(* IEC 61131-3 sources: avi-aoi-management/scripts/ai-eval/ngau-nhien/kho/st-ud5-sao-tam-giac/khung/src, 2 files *)

(* ---- KhoaChuyenMach.st ---- *)
FUNCTION_BLOCK KhoaChuyenMach
VAR_INPUT
    YC_SAO : BOOL;
    YC_TG : BOOL;
END_VAR
VAR_OUTPUT
    KM_SAO : BOOL;
    KM_TAM_GIAC : BOOL;
END_VAR
    (* TODO: cài đặt theo đề bài *)
    KM_SAO := FALSE;
END_FUNCTION_BLOCK

(* ---- KhoiDongSaoTamGiac.st ---- *)
FUNCTION_BLOCK KhoiDongSaoTamGiac
VAR_INPUT
    START : BOOL;
    STOP : BOOL;
    QUA_TAI : BOOL;
    RESET : BOOL;
    T_SAO : TIME;
    T_KHE : TIME;
END_VAR
VAR_OUTPUT
    KM_CHINH : BOOL;
    KM_SAO : BOOL;
    KM_TAM_GIAC : BOOL;
    LOI_QT : BOOL;
    TRANG_THAI : INT;
END_VAR
    (* TODO: cài đặt theo đề bài *)
    KM_CHINH := FALSE;
END_FUNCTION_BLOCK
